Fanuc KAREL source: KB00140.KL

PROGRAM KB00140
%NOLOCKGROUP
%ENVIRONMENT CORE
VAR
  P1: STRING[80]
  P2: INTEGER
BEGIN
  P1 = 'A'
  P2 = 1
  PROG_RESTORE(P1, P2)
END KB00140
